INTERFACE I_Diagnosable EXTENDS __SYSTEM.IQueryInterface

PROPERTY Name      : STRING
GET
END_GET
END_PROPERTY

PROPERTY HasFault  : BOOL
GET
END_GET
END_PROPERTY

PROPERTY FaultText : STRING
GET
END_GET
END_PROPERTY

END_INTERFACE

(* stored: Version 1.1.0.1
   Itf I_Diagnosable: Id {ccfd0e33-5c65-4a21-b2be-3f8a17641aa6}
   Property Name: Id {08ea8245-8117-4fe6-b074-011a233ea390}
   Get Get: Id {7b7478c0-50e3-40b2-9b2f-6539beaeb538}
   Property HasFault: Id {2e69767f-5e10-49f9-9e68-27d91c18d7c4}
   Get Get: Id {613758ed-47bf-453d-a772-8f43f9666d87}
   Property FaultText: Id {36eafa02-d8d1-4b06-bb84-d1aac5ebc7fe}
   Get Get: Id {bfc05c9f-fd9a-4ddb-9787-b3bc9a41b583} *)
